// Mitsubishi GX Works2 project: 金达路一号停车场洗车机   PLC: FX3U/FX3UC

PROGRAM MAIN
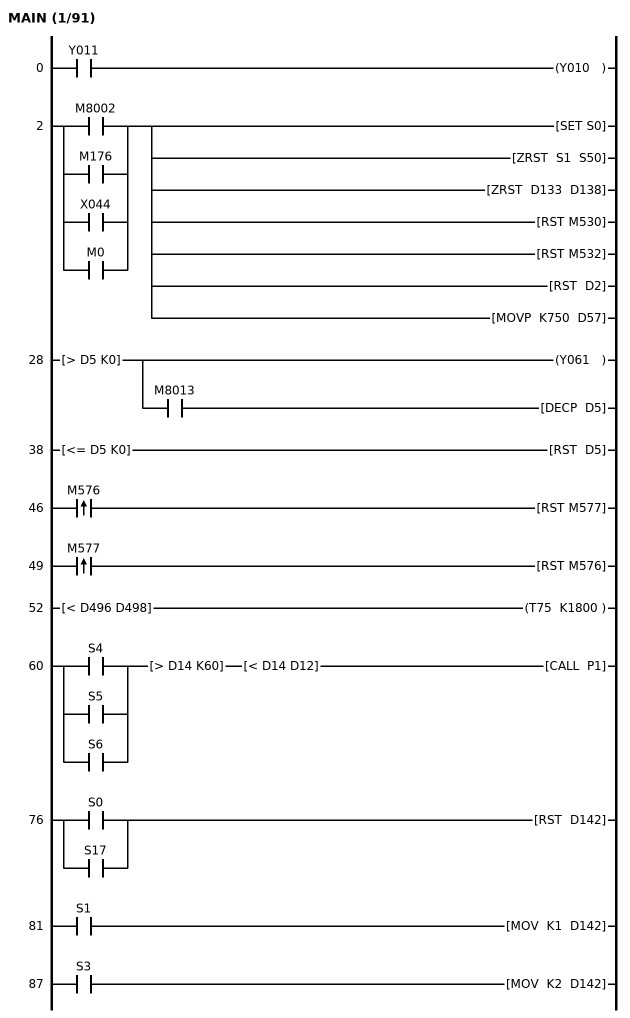
0     LD      Y011
      OUT     Y010
2     LD      M8002
      OR      M176
      OR      X044
      OR      M0
      SET     S0
      ZRST    S1 S50
      ZRST    D133 D138
      RST     M530
      RST     M532
      RST     D2
      MOVP    K750 D57
28    LD>     D5 K0
      OUT     Y061
      AND     M8013
      DECP    D5
38    LD<=    D5 K0
      RST     D5
46    LDP     M576
      RST     M577
49    LDP     M577
      RST     M576
52    LD<     D496 D498
      OUT     T75 K1800
60    LD      S4
      OR      S5
      OR      S6
      AND>    D14 K60
      AND<    D14 D12
      CALL    P1
76    LD      S0
      OR      S17
      RST     D142
81    LD      S1
      MOV     K1 D142
87    LD      S3
      MOV     K2 D142
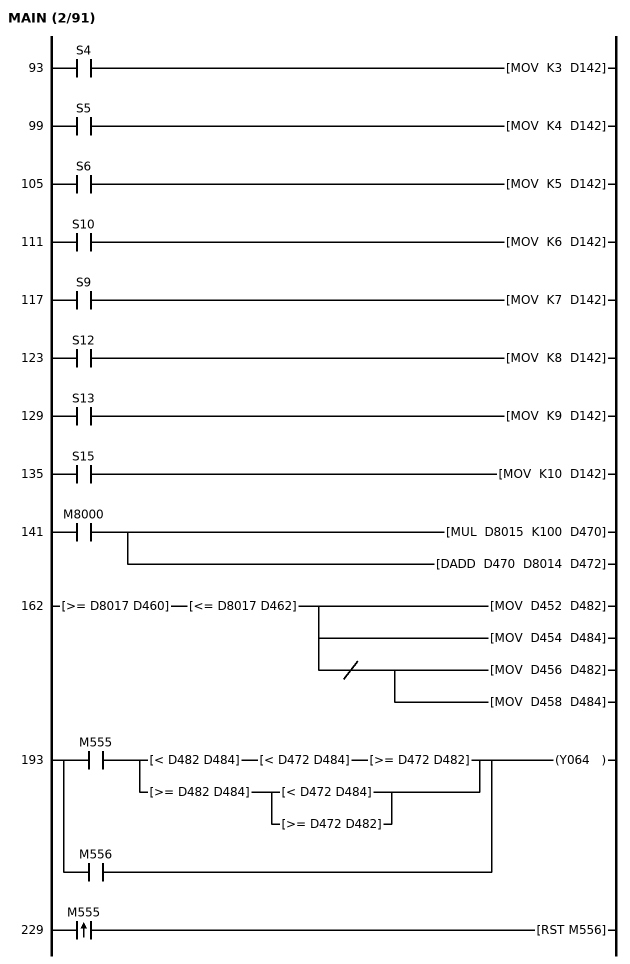
93    LD      S4
      MOV     K3 D142
99    LD      S5
      MOV     K4 D142
105   LD      S6
      MOV     K5 D142
111   LD      S10
      MOV     K6 D142
117   LD      S9
      MOV     K7 D142
123   LD      S12
      MOV     K8 D142
129   LD      S13
      MOV     K9 D142
135   LD      S15
      MOV     K10 D142
141   LD      M8000
      MUL     D8015 K100 D470
      DADD    D470 D8014 D472
162   LD>=    D8017 D460
      AND<=   D8017 D462
      MOV     D452 D482
      MOV     D454 D484
      INV
      MOV     D456 D482
      MOV     D458 D484
193   LD      M555
      LD<     D482 D484
      AND<    D472 D484
      AND>=   D472 D482
      LD>=    D482 D484
      LD<     D472 D484
      OR>=    D472 D482
      ANB
      ORB
      ANB
      OR      M556
      OUT     Y064
229   LDP     M555
      RST     M556
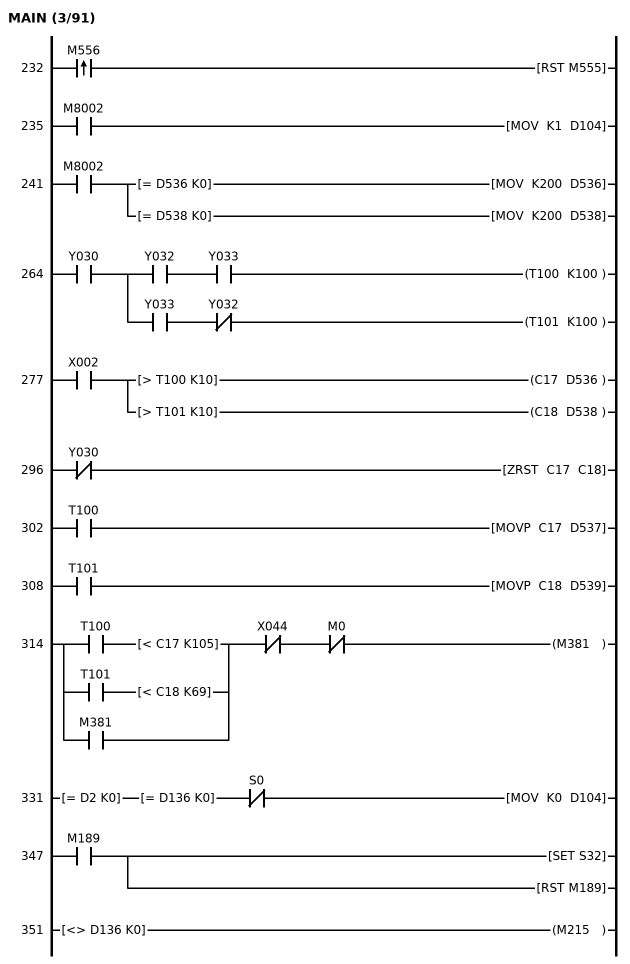
232   LDP     M556
      RST     M555
235   LD      M8002
      MOV     K1 D104
241   LD      M8002
      MPS
      AND=    D536 K0
      MOV     K200 D536
      MPP
      AND=    D538 K0
      MOV     K200 D538
264   LD      Y030
      MPS
      AND     Y032
      AND     Y033
      OUT     T100 K100
      MPP
      AND     Y033
      ANI     Y032
      OUT     T101 K100
277   LD      X002
      MPS
      AND>    T100 K10
      OUT     C17 D536
      MPP
      AND>    T101 K10
      OUT     C18 D538
296   LDI     Y030
      ZRST    C17 C18
302   LD      T100
      MOVP    C17 D537
308   LD      T101
      MOVP    C18 D539
314   LD      T100
      AND<    C17 K105
      LD      T101
      AND<    C18 K69
      ORB
      OR      M381
      ANI     X044
      ANI     M0
      OUT     M381
331   LD=     D2 K0
      AND=    D136 K0
      ANI     S0
      MOV     K0 D104
347   LD      M189
      SET     S32
      RST     M189
351   LD<>    D136 K0
      OUT     M215
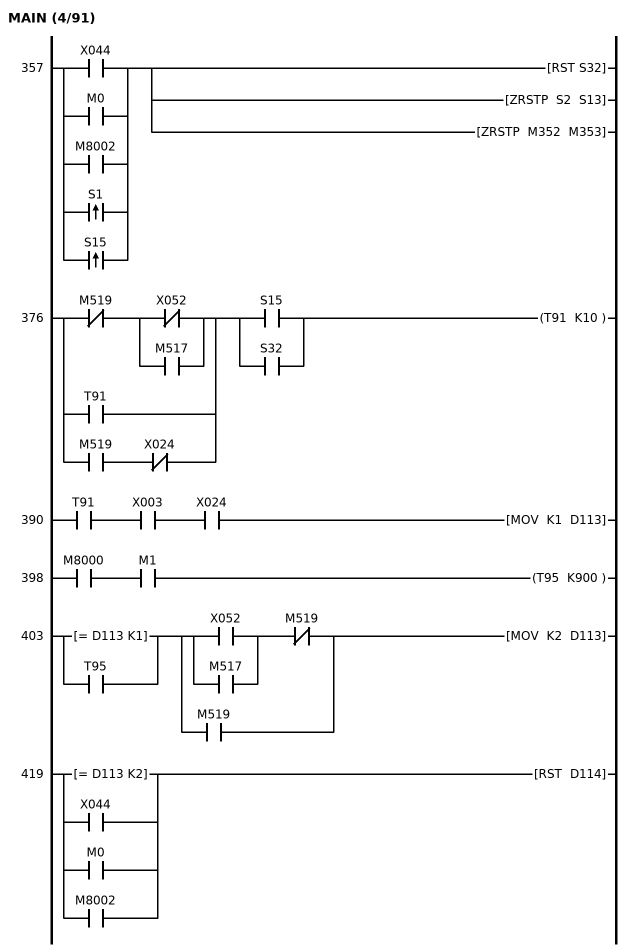
357   LD      X044
      OR      M0
      OR      M8002
      ORP     S1
      ORP     S15
      RST     S32
      ZRSTP   S2 S13
      ZRSTP   M352 M353
376   LDI     M519
      LDI     X052
      OR      M517
      ANB
      OR      T91
      LD      M519
      ANI     X024
      ORB
      LD      S15
      OR      S32
      ANB
      OUT     T91 K10
390   LD      T91
      AND     X003
      AND     X024
      MOV     K1 D113
398   LD      M8000
      AND     M1
      OUT     T95 K900
403   LD=     D113 K1
      OR      T95
      LD      X052
      OR      M517
      ANI     M519
      OR      M519
      ANB
      MOV     K2 D113
419   LD=     D113 K2
      OR      X044
      OR      M0
      OR      M8002
      RST     D114
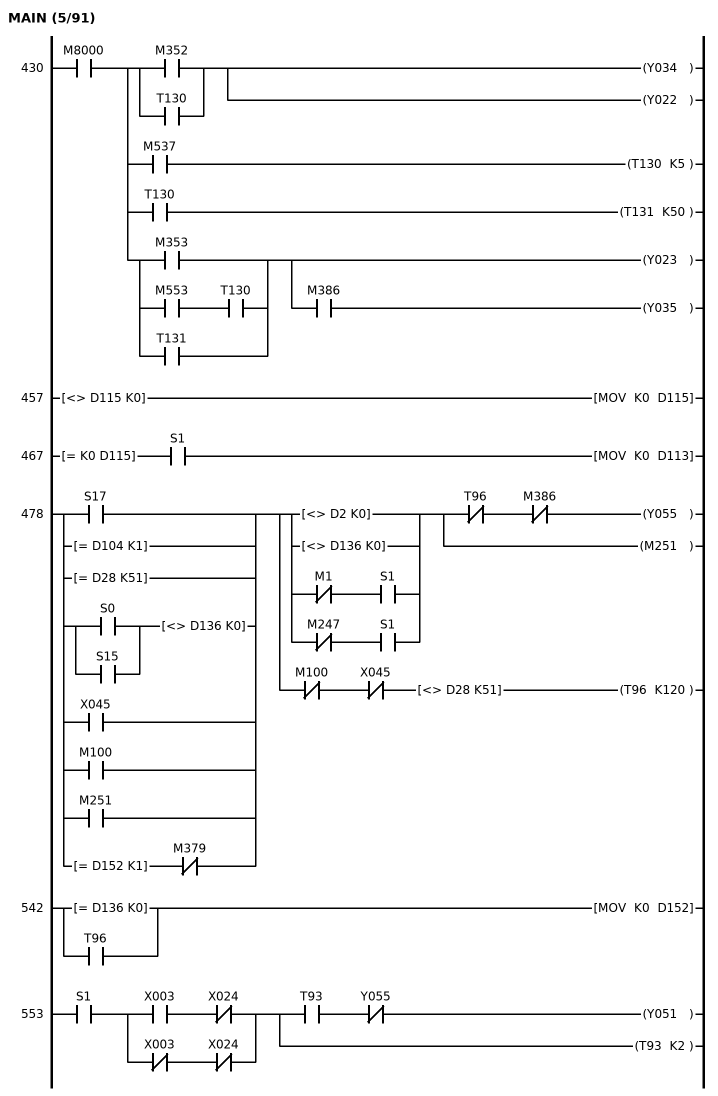
430   LD      M8000
      MPS
      LD      M352
      OR      T130
      ANB
      OUT     Y034
      OUT     Y022
      MRD
      AND     M537
      OUT     T130 K5
      MRD
      AND     T130
      OUT     T131 K50
      MPP
      LD      M353
      LD      M553
      AND     T130
      ORB
      OR      T131
      ANB
      OUT     Y023
      AND     M386
      OUT     Y035
457   LD<>    D115 K0
      MOV     K0 D115
467   LD=     K0 D115
      AND     S1
      MOV     K0 D113
478   LD      S17
      OR=     D104 K1
      OR=     D28 K51
      LD      S0
      OR      S15
      AND<>   D136 K0
      ORB
      OR      X045
      OR      M100
      OR      M251
      LD=     D152 K1
      ANI     M379
      ORB
      MPS
      LD<>    D2 K0
      OR<>    D136 K0
      LDI     M1
      AND     S1
      ORB
      LDI     M247
      AND     S1
      ORB
      ANB
      MPS
      ANI     T96
      ANI     M386
      OUT     Y055
      MPP
      OUT     M251
      MPP
      ANI     M100
      ANI     X045
      AND<>   D28 K51
      OUT     T96 K120
542   LD=     D136 K0
      OR      T96
      MOV     K0 D152
553   LD      S1
      LD      X003
      ANI     X024
      LDI     X003
      ANI     X024
      ORB
      ANB
      MPS
      AND     T93
      ANI     Y055
      OUT     Y051
      MPP
      OUT     T93 K2
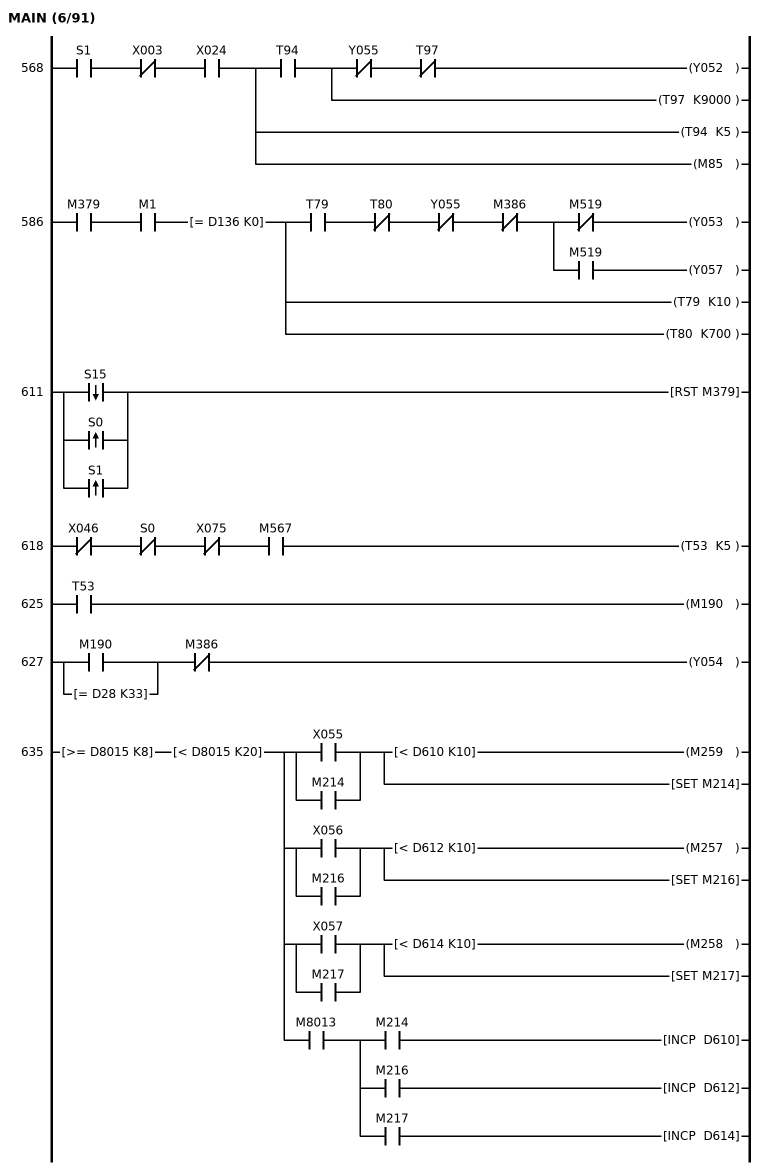
568   LD      S1
      ANI     X003
      AND     X024
      MPS
      AND     T94
      MPS
      ANI     Y055
      ANI     T97
      OUT     Y052
      MPP
      OUT     T97 K9000
      MPP
      OUT     T94 K5
      OUT     M85
586   LD      M379
      AND     M1
      AND=    D136 K0
      MPS
      AND     T79
      ANI     T80
      ANI     Y055
      ANI     M386
      MPS
      ANI     M519
      OUT     Y053
      MPP
      AND     M519
      OUT     Y057
      MPP
      OUT     T79 K10
      OUT     T80 K700
611   LDF     S15
      ORP     S0
      ORP     S1
      RST     M379
618   LDI     X046
      ANI     S0
      ANI     X075
      AND     M567
      OUT     T53 K5
625   LD      T53
      OUT     M190
627   LD      M190
      OR=     D28 K33
      ANI     M386
      OUT     Y054
635   LD>=    D8015 K8
      AND<    D8015 K20
      MPS
      LD      X055
      OR      M214
      ANB
      MPS
      AND<    D610 K10
      OUT     M259
      MPP
      SET     M214
      MRD
      LD      X056
      OR      M216
      ANB
      MPS
      AND<    D612 K10
      OUT     M257
      MPP
      SET     M216
      MRD
      LD      X057
      OR      M217
      ANB
      MPS
      AND<    D614 K10
      OUT     M258
      MPP
      SET     M217
      MPP
      AND     M8013
      MPS
      AND     M214
      INCP    D610
      MRD
      AND     M216
      INCP    D612
      MPP
      AND     M217
      INCP    D614
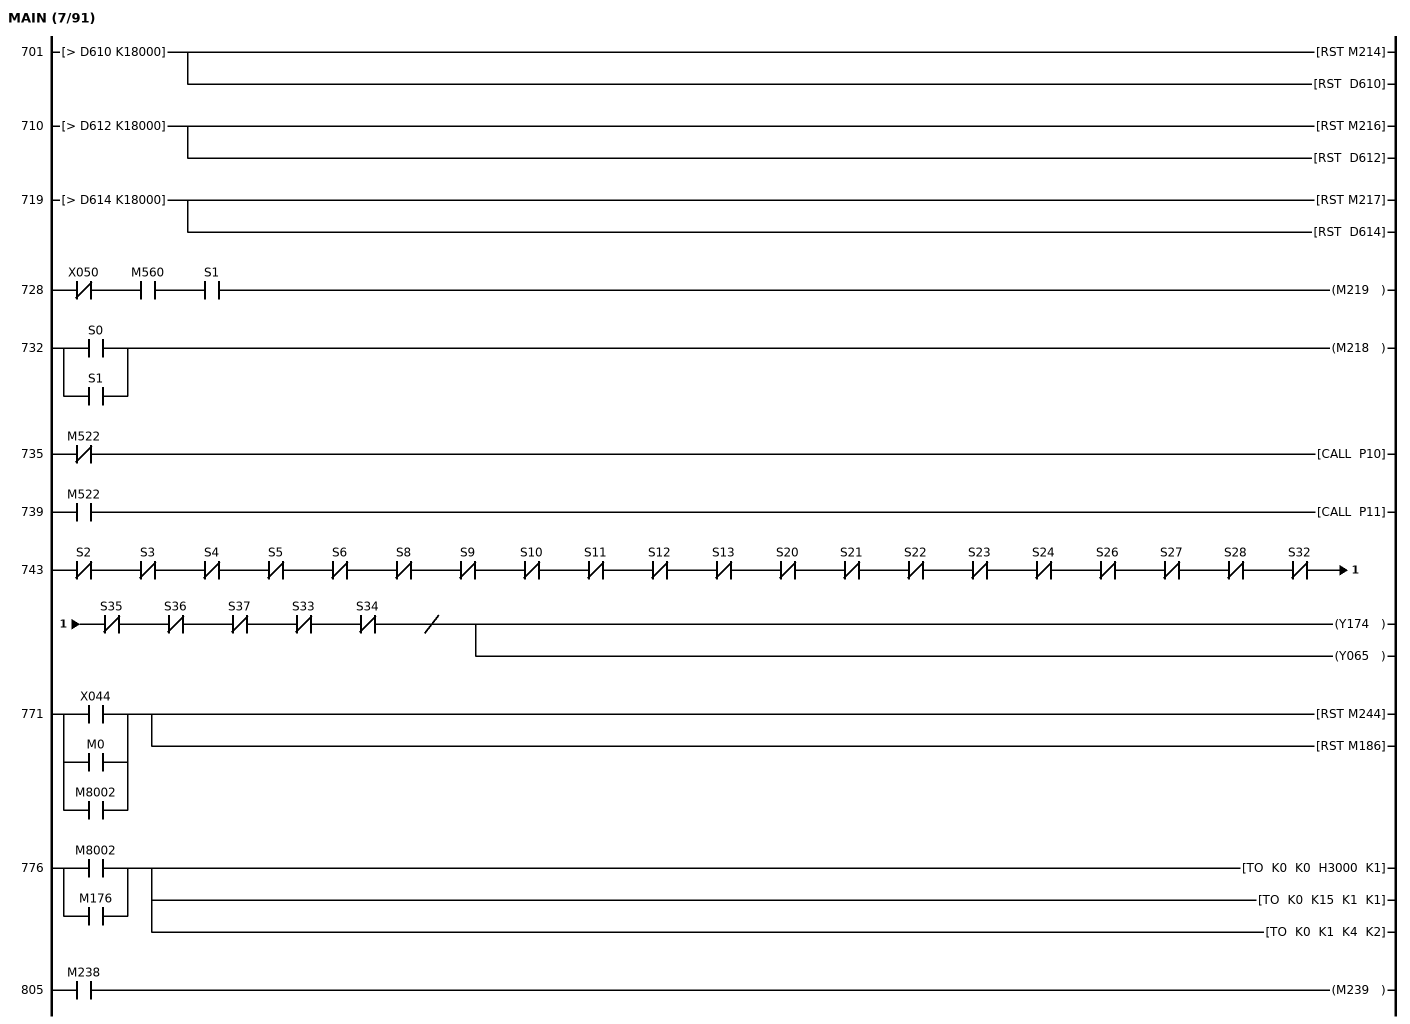
701   LD>     D610 K18000
      RST     M214
      RST     D610
710   LD>     D612 K18000
      RST     M216
      RST     D612
719   LD>     D614 K18000
      RST     M217
      RST     D614
728   LDI     X050
      AND     M560
      AND     S1
      OUT     M219
732   LD      S0
      OR      S1
      OUT     M218
735   LDI     M522
      CALL    P10
739   LD      M522
      CALL    P11
743   LDI     S2
      ANI     S3
      ANI     S4
      ANI     S5
      ANI     S6
      ANI     S8
      ANI     S9
      ANI     S10
      ANI     S11
      ANI     S12
      ANI     S13
      ANI     S20
      ANI     S21
      ANI     S22
      ANI     S23
      ANI     S24
      ANI     S26
      ANI     S27
      ANI     S28
      ANI     S32
      ANI     S35
      ANI     S36
      ANI     S37
      ANI     S33
      ANI     S34
      INV
      OUT     Y174
      OUT     Y065
771   LD      X044
      OR      M0
      OR      M8002
      RST     M244
      RST     M186
776   LD      M8002
      OR      M176
      TO      K0 K0 H3000 K1
      TO      K0 K15 K1 K1
      TO      K0 K1 K4 K2
805   LD      M238
      OUT     M239
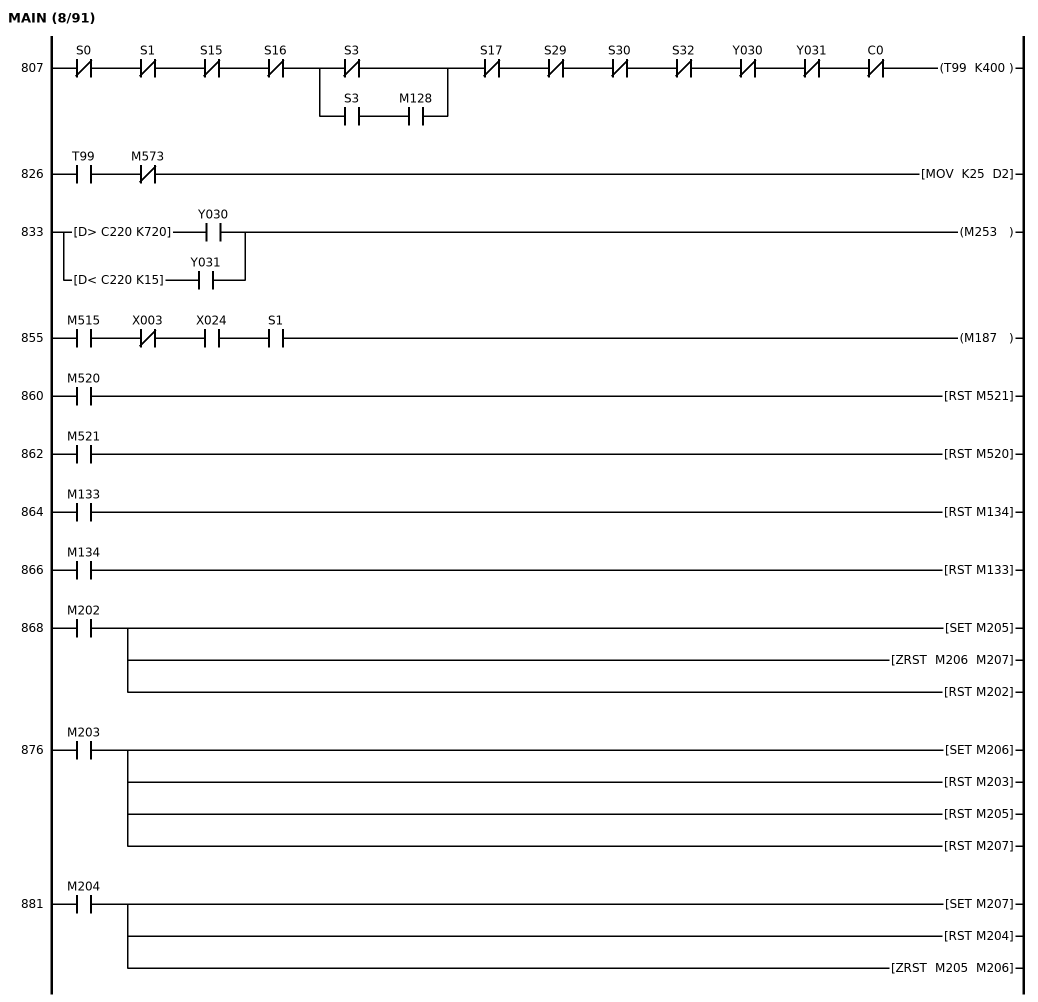
807   LDI     S0
      ANI     S1
      ANI     S15
      ANI     S16
      LDI     S3
      LD      S3
      AND     M128
      ORB
      ANB
      ANI     S17
      ANI     S29
      ANI     S30
      ANI     S32
      ANI     Y030
      ANI     Y031
      ANI     C0
      OUT     T99 K400
826   LD      T99
      ANI     M573
      MOV     K25 D2
833   LDD>    C220 K720
      AND     Y030
      LDD<    C220 K15
      AND     Y031
      ORB
      OUT     M253
855   LD      M515
      ANI     X003
      AND     X024
      AND     S1
      OUT     M187
860   LD      M520
      RST     M521
862   LD      M521
      RST     M520
864   LD      M133
      RST     M134
866   LD      M134
      RST     M133
868   LD      M202
      SET     M205
      ZRST    M206 M207
      RST     M202
876   LD      M203
      SET     M206
      RST     M203
      RST     M205
      RST     M207
881   LD      M204
      SET     M207
      RST     M204
      ZRST    M205 M206
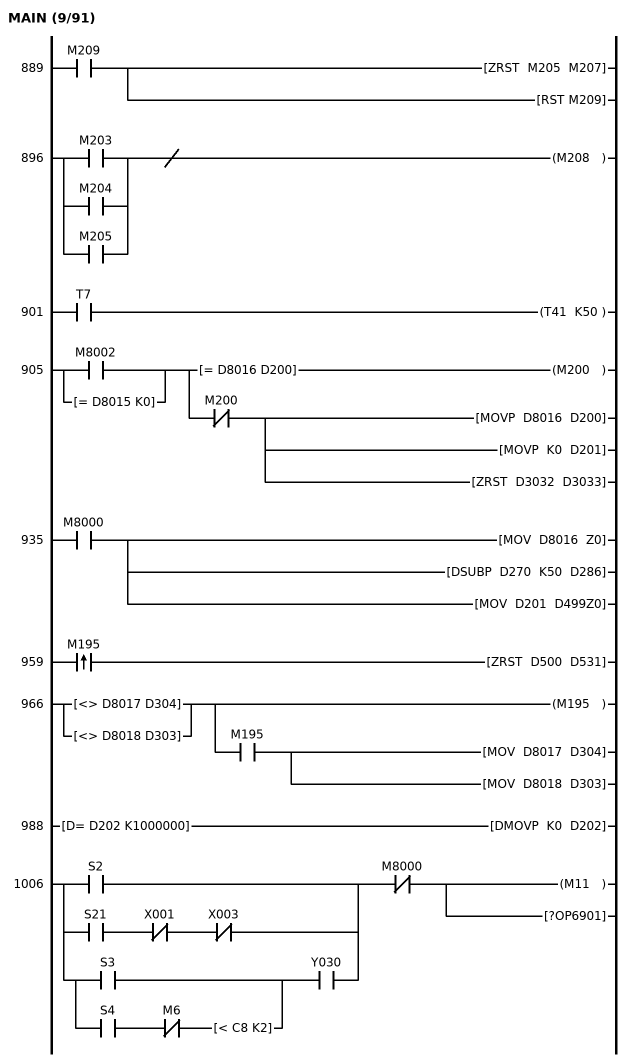
889   LD      M209
      ZRST    M205 M207
      RST     M209
896   LD      M203
      OR      M204
      OR      M205
      INV
      OUT     M208
901   LD      T7
      OUT     T41 K50
905   LD      M8002
      OR=     D8015 K0
      MPS
      AND=    D8016 D200
      OUT     M200
      MPP
      ANI     M200
      MOVP    D8016 D200
      MOVP    K0 D201
      ZRST    D3032 D3033
935   LD      M8000
      MOV     D8016 Z0
      DSUBP   D270 K50 D286
      MOV     D201 D499Z0
959   LDP     M195
      ZRST    D500 D531
966   LD<>    D8017 D304
      OR<>    D8018 D303
      OUT     M195
      AND     M195
      MOV     D8017 D304
      MOV     D8018 D303
988   LDD=    D202 K1000000
      DMOVP   K0 D202
1006  LD      S2
      LD      S21
      ANI     X001
      ANI     X003
      ORB
      LD      S3
      LD      S4
      ANI     M6
      AND<    C8 K2
      ORB
      AND     Y030
      ORB
      ANI     M8000
      OUT     M11
      ?OP6901
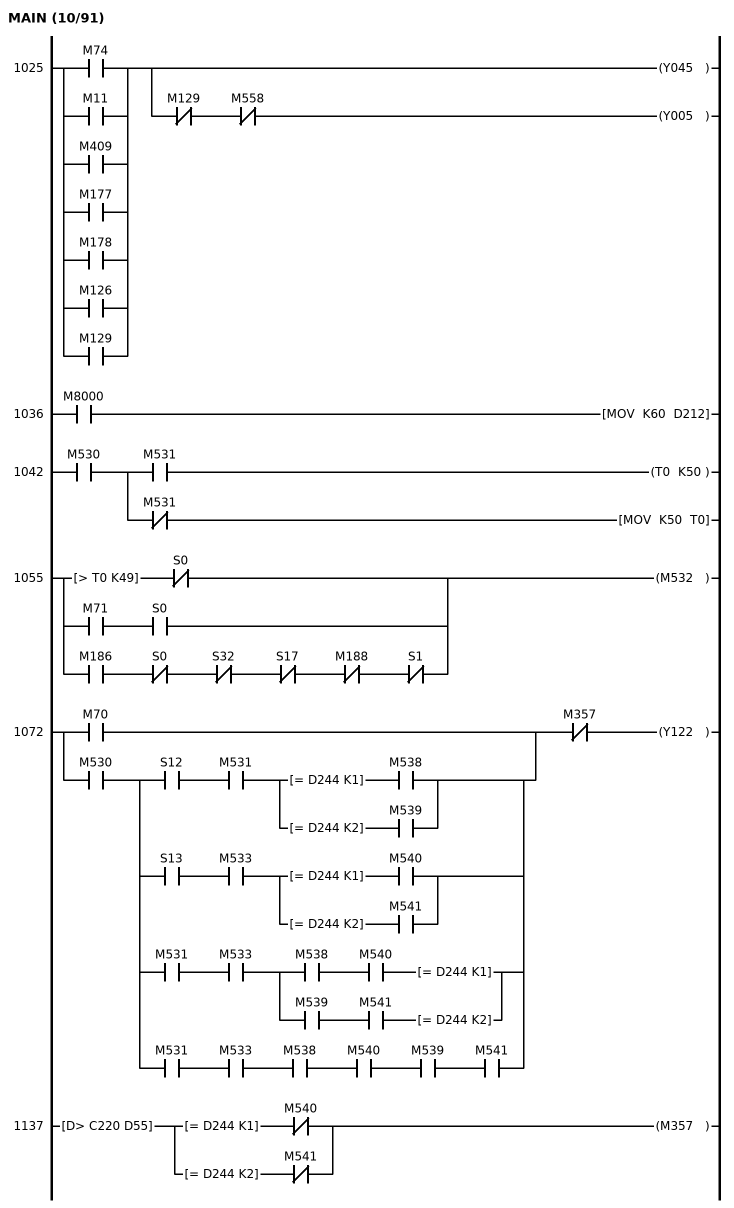
1025  LD      M74
      OR      M11
      OR      M409
      OR      M177
      OR      M178
      OR      M126
      OR      M129
      OUT     Y045
      ANI     M129
      ANI     M558
      OUT     Y005
1036  LD      M8000
      MOV     K60 D212
1042  LD      M530
      MPS
      AND     M531
      OUT     T0 K50
      MPP
      ANI     M531
      MOV     K50 T0
1055  LD>     T0 K49
      ANI     S0
      LD      M71
      AND     S0
      ORB
      LD      M186
      ANI     S0
      ANI     S32
      ANI     S17
      ANI     M188
      ANI     S1
      ORB
      OUT     M532
1072  LD      M70
      LD      M530
      LD      S12
      AND     M531
      LD=     D244 K1
      AND     M538
      LD=     D244 K2
      AND     M539
      ORB
      ANB
      LD      S13
      AND     M533
      LD=     D244 K1
      AND     M540
      LD=     D244 K2
      AND     M541
      ORB
      ANB
      ORB
      LD      M531
      AND     M533
      LD      M538
      AND     M540
      AND=    D244 K1
      LD      M539
      AND     M541
      AND=    D244 K2
      ORB
      ANB
      ORB
      LD      M531
      AND     M533
      AND     M538
      AND     M540
      AND     M539
      AND     M541
      ORB
      ANB
      ORB
      ANI     M357
      OUT     Y122
1137  LDD>    C220 D55
      LD=     D244 K1
      ANI     M540
      LD=     D244 K2
      ANI     M541
      ORB
      ANB
      OUT     M357
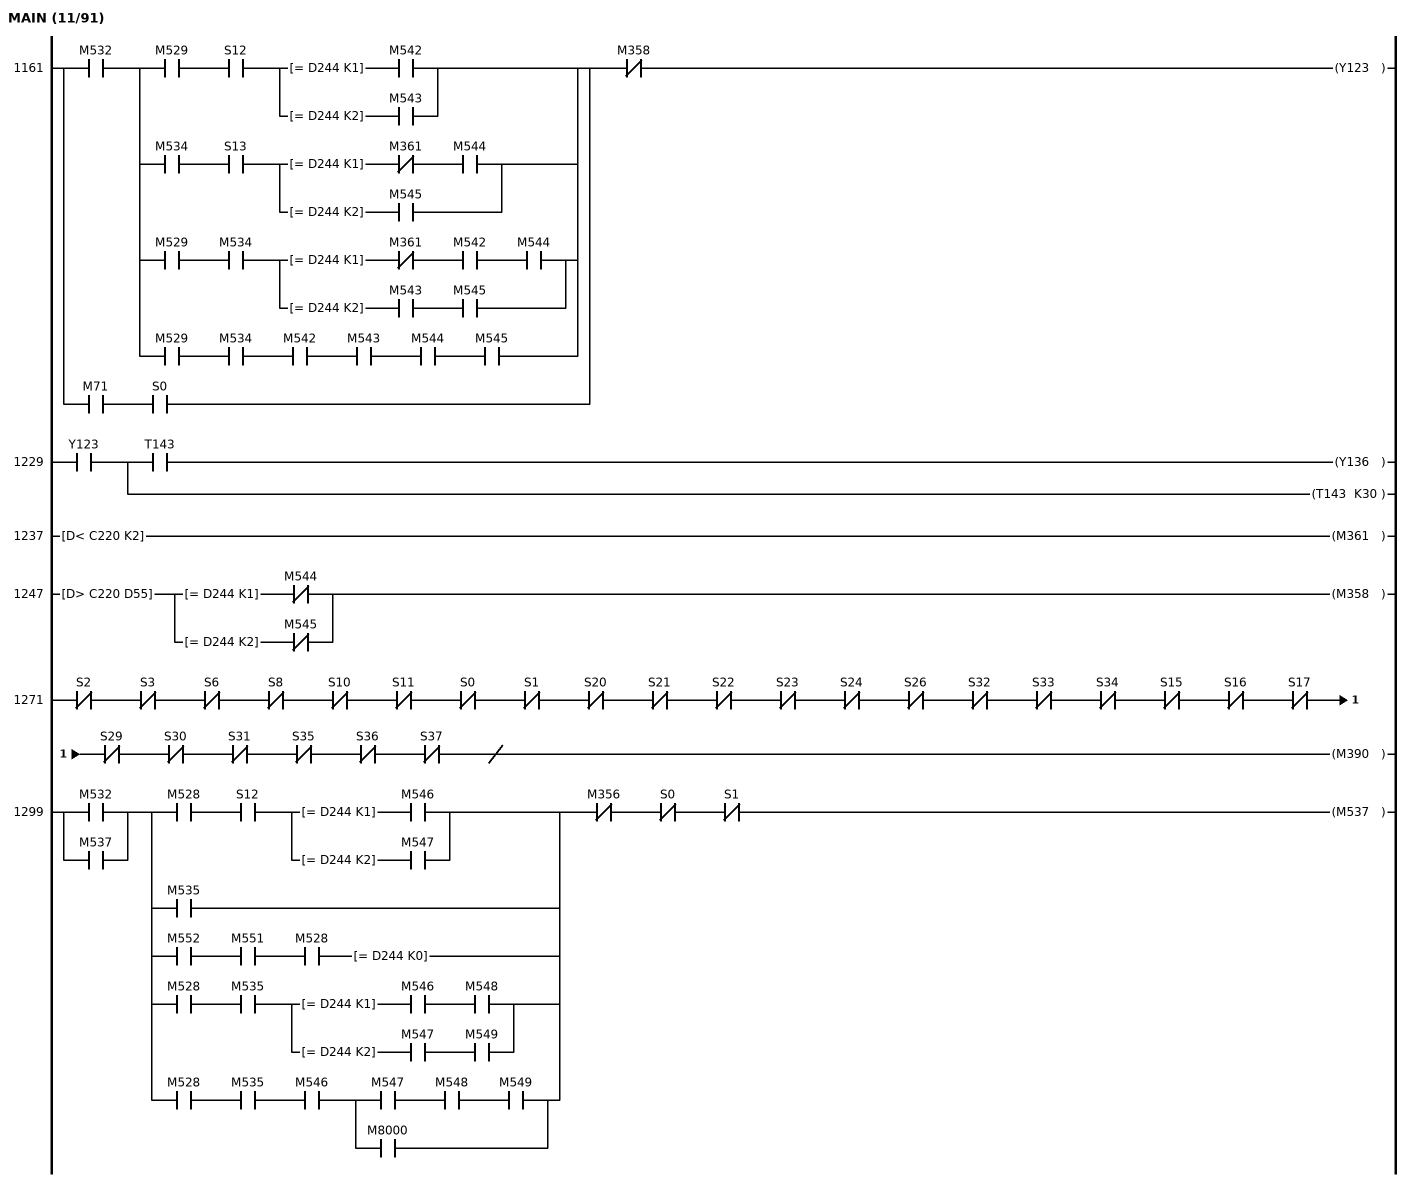
1161  LD      M532
      LD      M529
      AND     S12
      LD=     D244 K1
      AND     M542
      LD=     D244 K2
      AND     M543
      ORB
      ANB
      LD      M534
      AND     S13
      LD=     D244 K1
      ANI     M361
      AND     M544
      LD=     D244 K2
      AND     M545
      ORB
      ANB
      ORB
      LD      M529
      AND     M534
      LD=     D244 K1
      ANI     M361
      AND     M542
      AND     M544
      LD=     D244 K2
      AND     M543
      AND     M545
      ORB
      ANB
      ORB
      LD      M529
      AND     M534
      AND     M542
      AND     M543
      AND     M544
      AND     M545
      ORB
      ANB
      LD      M71
      AND     S0
      ORB
      ANI     M358
      OUT     Y123
1229  LD      Y123
      MPS
      AND     T143
      OUT     Y136
      MPP
      OUT     T143 K30
1237  LDD<    C220 K2
      OUT     M361
1247  LDD>    C220 D55
      LD=     D244 K1
      ANI     M544
      LD=     D244 K2
      ANI     M545
      ORB
      ANB
      OUT     M358
1271  LDI     S2
      ANI     S3
      ANI     S6
      ANI     S8
      ANI     S10
      ANI     S11
      ANI     S0
      ANI     S1
      ANI     S20
      ANI     S21
      ANI     S22
      ANI     S23
      ANI     S24
      ANI     S26
      ANI     S32
      ANI     S33
      ANI     S34
      ANI     S15
      ANI     S16
      ANI     S17
      ANI     S29
      ANI     S30
      ANI     S31
      ANI     S35
      ANI     S36
      ANI     S37
      INV
      OUT     M390
1299  LD      M532
      OR      M537
      LD      M528
      AND     S12
      LD=     D244 K1
      AND     M546
      LD=     D244 K2
      AND     M547
      ORB
      ANB
      OR      M535
      LD      M552
      AND     M551
      AND     M528
      AND=    D244 K0
      ORB
      LD      M528
      AND     M535
      LD=     D244 K1
      AND     M546
      AND     M548
      LD=     D244 K2
      AND     M547
      AND     M549
      ORB
      ANB
      ORB
      LD      M528
      AND     M535
      AND     M546
      LD      M547
      AND     M548
      AND     M549
      OR      M8000
      ANB
      ORB
      ANB
      ANI     M356
      ANI     S0
      ANI     S1
      OUT     M537
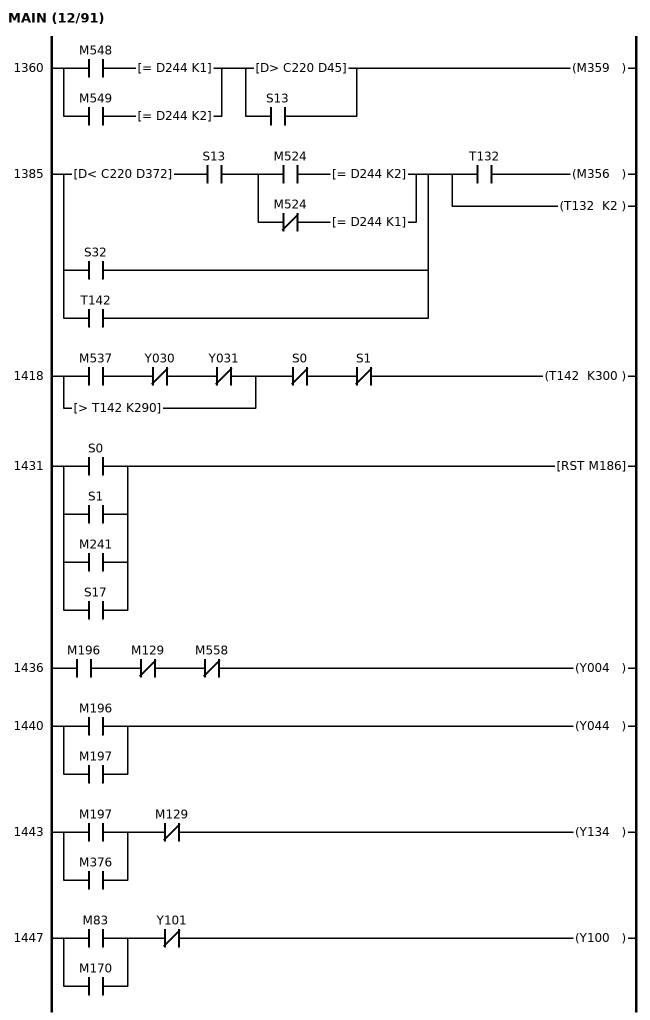
1360  LD      M548
      AND=    D244 K1
      LD      M549
      AND=    D244 K2
      ORB
      LDD>    C220 D45
      OR      S13
      ANB
      OUT     M359
1385  LDD<    C220 D372
      AND     S13
      LD      M524
      AND=    D244 K2
      LDI     M524
      AND=    D244 K1
      ORB
      ANB
      OR      S32
      OR      T142
      MPS
      AND     T132
      OUT     M356
      MPP
      OUT     T132 K2
1418  LD      M537
      ANI     Y030
      ANI     Y031
      OR>     T142 K290
      ANI     S0
      ANI     S1
      OUT     T142 K300
1431  LD      S0
      OR      S1
      OR      M241
      OR      S17
      RST     M186
1436  LD      M196
      ANI     M129
      ANI     M558
      OUT     Y004
1440  LD      M196
      OR      M197
      OUT     Y044
1443  LD      M197
      OR      M376
      ANI     M129
      OUT     Y134
1447  LD      M83
      OR      M170
      ANI     Y101
      OUT     Y100
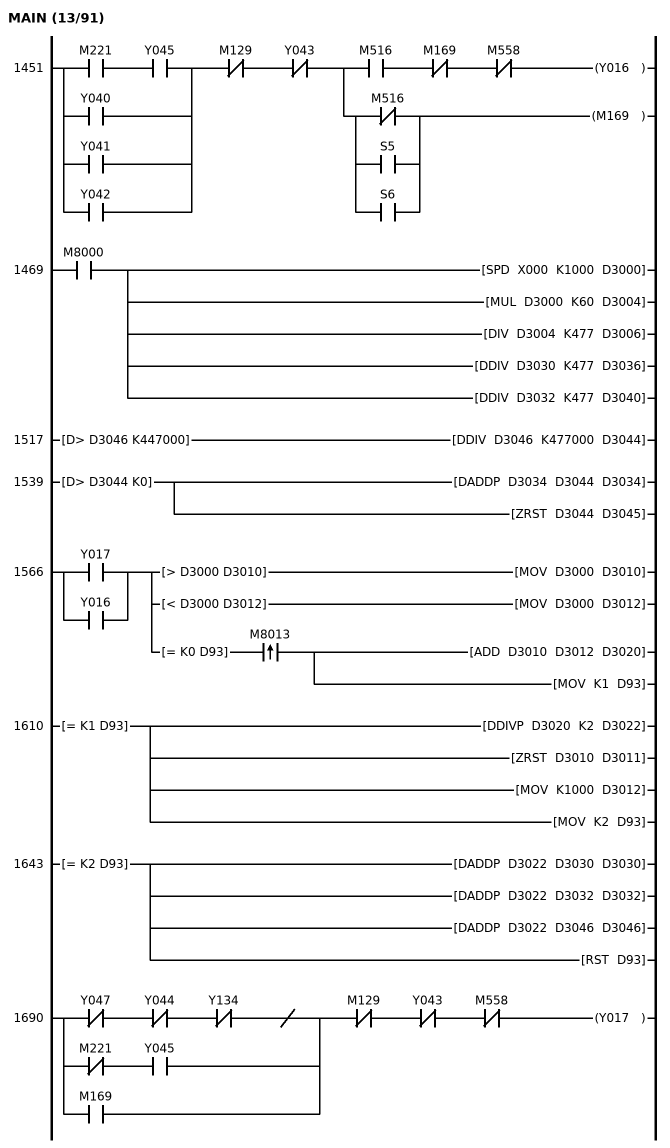
1451  LD      M221
      AND     Y045
      OR      Y040
      OR      Y041
      OR      Y042
      ANI     M129
      ANI     Y043
      MPS
      AND     M516
      ANI     M169
      ANI     M558
      OUT     Y016
      MPP
      LDI     M516
      OR      S5
      OR      S6
      ANB
      OUT     M169
1469  LD      M8000
      SPD     X000 K1000 D3000
      MUL     D3000 K60 D3004
      DIV     D3004 K477 D3006
      DDIV    D3030 K477 D3036
      DDIV    D3032 K477 D3040
1517  LDD>    D3046 K447000
      DDIV    D3046 K477000 D3044
1539  LDD>    D3044 K0
      DADDP   D3034 D3044 D3034
      ZRST    D3044 D3045
1566  LD      Y017
      OR      Y016
      MPS
      AND>    D3000 D3010
      MOV     D3000 D3010
      MRD
      AND<    D3000 D3012
      MOV     D3000 D3012
      MPP
      AND=    K0 D93
      ANDP    M8013
      ADD     D3010 D3012 D3020
      MOV     K1 D93
1610  LD=     K1 D93
      DDIVP   D3020 K2 D3022
      ZRST    D3010 D3011
      MOV     K1000 D3012
      MOV     K2 D93
1643  LD=     K2 D93
      DADDP   D3022 D3030 D3030
      DADDP   D3022 D3032 D3032
      DADDP   D3022 D3046 D3046
      RST     D93
1690  LDI     Y047
      ANI     Y044
      ANI     Y134
      INV
      LDI     M221
      AND     Y045
      ORB
      OR      M169
      ANI     M129
      ANI     Y043
      ANI     M558
      OUT     Y017
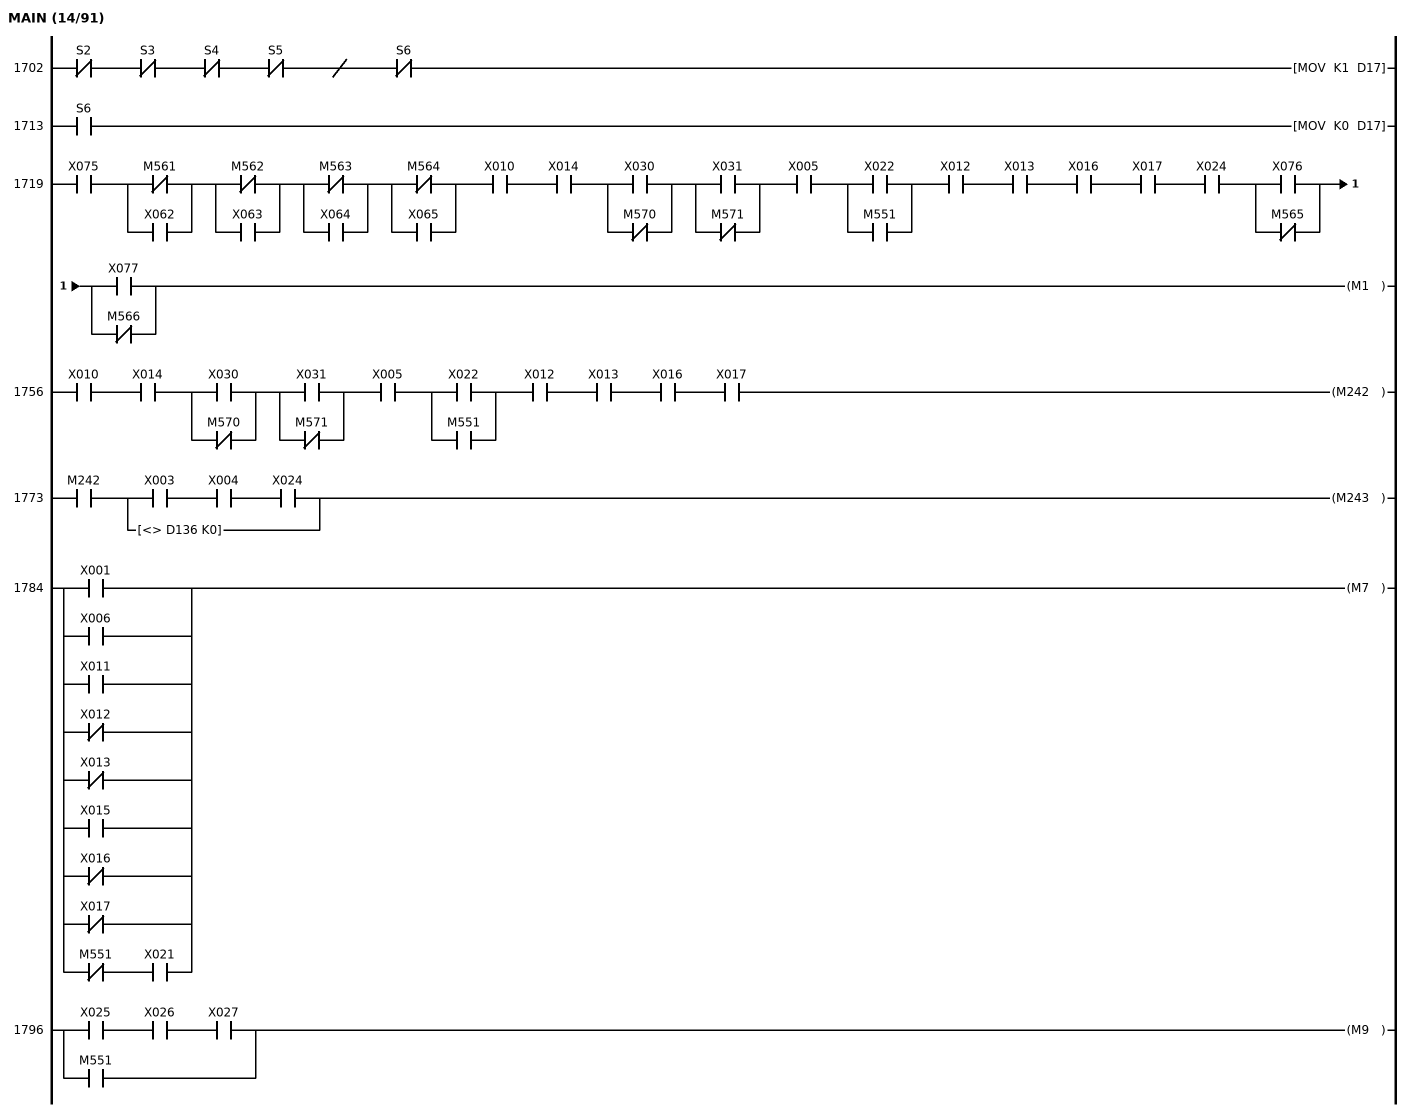
1702  LDI     S2
      ANI     S3
      ANI     S4
      ANI     S5
      INV
      ANI     S6
      MOV     K1 D17
1713  LD      S6
      MOV     K0 D17
1719  LD      X075
      LDI     M561
      OR      X062
      ANB
      LDI     M562
      OR      X063
      ANB
      LDI     M563
      OR      X064
      ANB
      LDI     M564
      OR      X065
      ANB
      AND     X010
      AND     X014
      LD      X030
      ORI     M570
      ANB
      LD      X031
      ORI     M571
      ANB
      AND     X005
      LD      X022
      OR      M551
      ANB
      AND     X012
      AND     X013
      AND     X016
      AND     X017
      AND     X024
      LD      X076
      ORI     M565
      ANB
      LD      X077
      ORI     M566
      ANB
      OUT     M1
1756  LD      X010
      AND     X014
      LD      X030
      ORI     M570
      ANB
      LD      X031
      ORI     M571
      ANB
      AND     X005
      LD      X022
      OR      M551
      ANB
      AND     X012
      AND     X013
      AND     X016
      AND     X017
      OUT     M242
1773  LD      M242
      LD      X003
      AND     X004
      AND     X024
      OR<>    D136 K0
      ANB
      OUT     M243
1784  LD      X001
      OR      X006
      OR      X011
      ORI     X012
      ORI     X013
      OR      X015
      ORI     X016
      ORI     X017
      LDI     M551
      AND     X021
      ORB
      OUT     M7
1796  LD      X025
      AND     X026
      AND     X027
      OR      M551
      OUT     M9
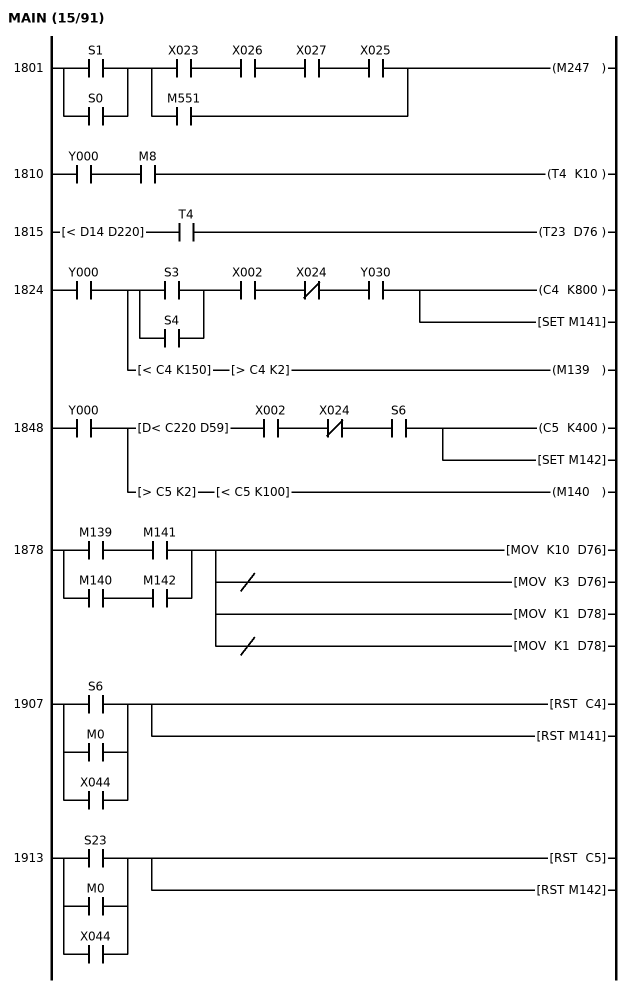
1801  LD      S1
      OR      S0
      LD      X023
      AND     X026
      AND     X027
      AND     X025
      OR      M551
      ANB
      OUT     M247
1810  LD      Y000
      AND     M8
      OUT     T4 K10
1815  LD<     D14 D220
      AND     T4
      OUT     T23 D76
1824  LD      Y000
      MPS
      LD      S3
      OR      S4
      ANB
      AND     X002
      ANI     X024
      AND     Y030
      OUT     C4 K800
      SET     M141
      MPP
      AND<    C4 K150
      AND>    C4 K2
      OUT     M139
1848  LD      Y000
      MPS
      ANDD<   C220 D59
      AND     X002
      ANI     X024
      AND     S6
      OUT     C5 K400
      SET     M142
      MPP
      AND>    C5 K2
      AND<    C5 K100
      OUT     M140
1878  LD      M139
      AND     M141
      LD      M140
      AND     M142
      ORB
      MOV     K10 D76
      MPS
      INV
      MOV     K3 D76
      MPP
      MOV     K1 D78
      INV
      MOV     K1 D78
1907  LD      S6
      OR      M0
      OR      X044
      RST     C4
      RST     M141
1913  LD      S23
      OR      M0
      OR      X044
      RST     C5
      RST     M142
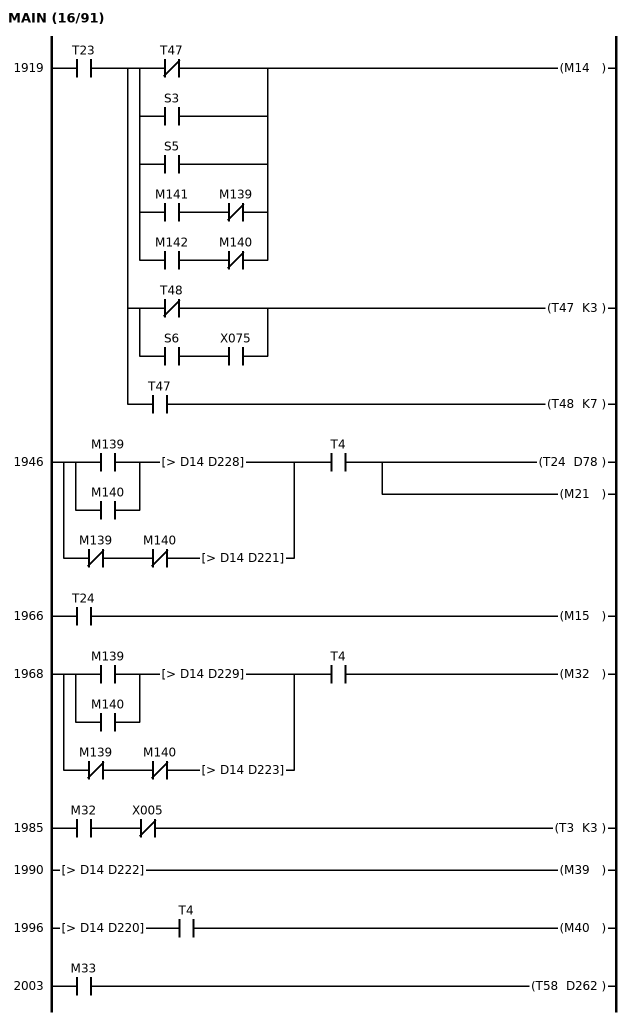
1919  LD      T23
      MPS
      LDI     T47
      OR      S3
      OR      S5
      LD      M141
      ANI     M139
      ORB
      LD      M142
      ANI     M140
      ORB
      ANB
      OUT     M14
      MRD
      LDI     T48
      LD      S6
      AND     X075
      ORB
      ANB
      OUT     T47 K3
      MPP
      AND     T47
      OUT     T48 K7
1946  LD      M139
      OR      M140
      AND>    D14 D228
      LDI     M139
      ANI     M140
      AND>    D14 D221
      ORB
      AND     T4
      OUT     T24 D78
      OUT     M21
1966  LD      T24
      OUT     M15
1968  LD      M139
      OR      M140
      AND>    D14 D229
      LDI     M139
      ANI     M140
      AND>    D14 D223
      ORB
      AND     T4
      OUT     M32
1985  LD      M32
      ANI     X005
      OUT     T3 K3
1990  LD>     D14 D222
      OUT     M39
1996  LD>     D14 D220
      AND     T4
      OUT     M40
2003  LD      M33
      OUT     T58 D262
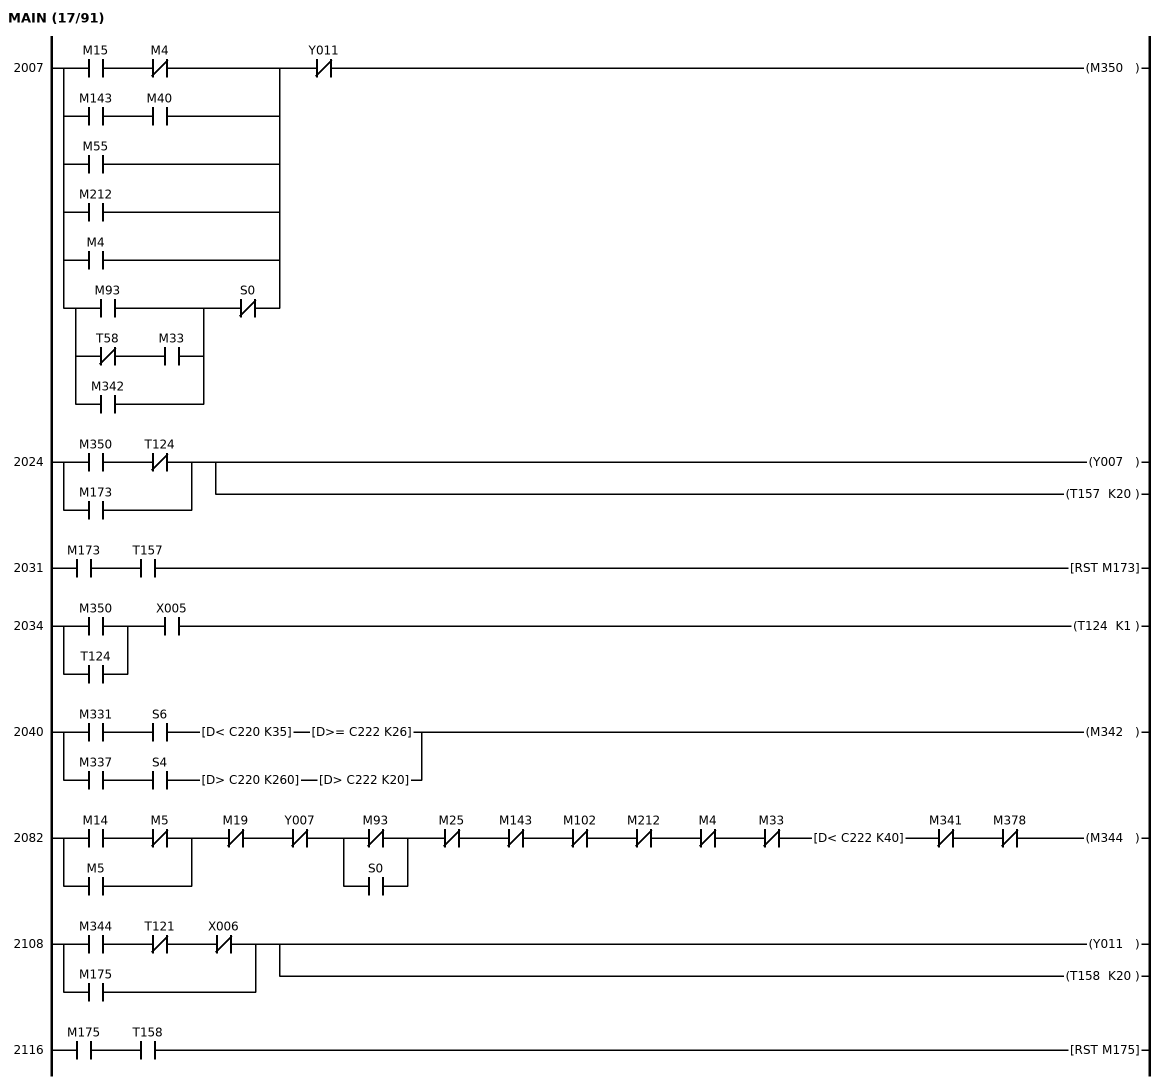
2007  LD      M15
      ANI     M4
      LD      M143
      AND     M40
      ORB
      OR      M55
      OR      M212
      OR      M4
      LD      M93
      LDI     T58
      AND     M33
      ORB
      OR      M342
      ANI     S0
      ORB
      ANI     Y011
      OUT     M350
2024  LD      M350
      ANI     T124
      OR      M173
      OUT     Y007
      OUT     T157 K20
2031  LD      M173
      AND     T157
      RST     M173
2034  LD      M350
      OR      T124
      AND     X005
      OUT     T124 K1
2040  LD      M331
      AND     S6
      ANDD<   C220 K35
      ANDD>=  C222 K26
      LD      M337
      AND     S4
      ANDD>   C220 K260
      ANDD>   C222 K20
      ORB
      OUT     M342
2082  LD      M14
      ANI     M5
      OR      M5
      ANI     M19
      ANI     Y007
      LDI     M93
      OR      S0
      ANB
      ANI     M25
      ANI     M143
      ANI     M102
      ANI     M212
      ANI     M4
      ANI     M33
      ANDD<   C222 K40
      ANI     M341
      ANI     M378
      OUT     M344
2108  LD      M344
      ANI     T121
      ANI     X006
      OR      M175
      OUT     Y011
      OUT     T158 K20
2116  LD      M175
      AND     T158
      RST     M175
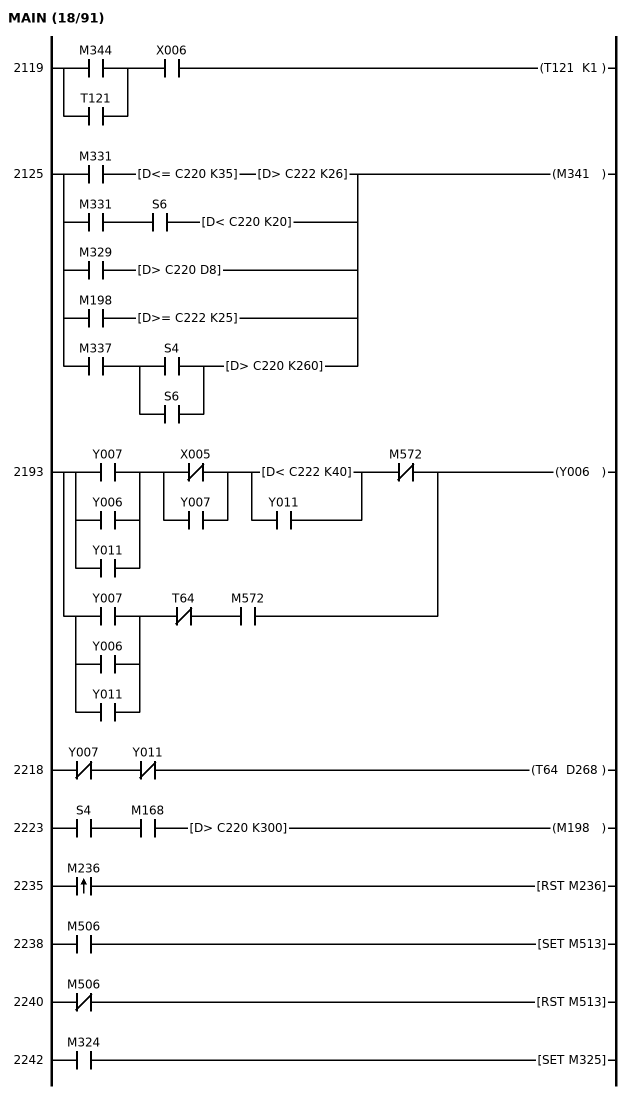
2119  LD      M344
      OR      T121
      AND     X006
      OUT     T121 K1
2125  LD      M331
      ANDD<=  C220 K35
      ANDD>   C222 K26
      LD      M331
      AND     S6
      ANDD<   C220 K20
      ORB
      LD      M329
      ANDD>   C220 D8
      ORB
      LD      M198
      ANDD>=  C222 K25
      ORB
      LD      M337
      LD      S4
      OR      S6
      ANB
      ANDD>   C220 K260
      ORB
      OUT     M341
2193  LD      Y007
      OR      Y006
      OR      Y011
      LDI     X005
      OR      Y007
      ANB
      LDD<    C222 K40
      OR      Y011
      ANB
      ANI     M572
      LD      Y007
      OR      Y006
      OR      Y011
      ANI     T64
      AND     M572
      ORB
      OUT     Y006
2218  LDI     Y007
      ANI     Y011
      OUT     T64 D268
2223  LD      S4
      AND     M168
      ANDD>   C220 K300
      OUT     M198
2235  LDP     M236
      RST     M236
2238  LD      M506
      SET     M513
2240  LDI     M506
      RST     M513
2242  LD      M324
      SET     M325
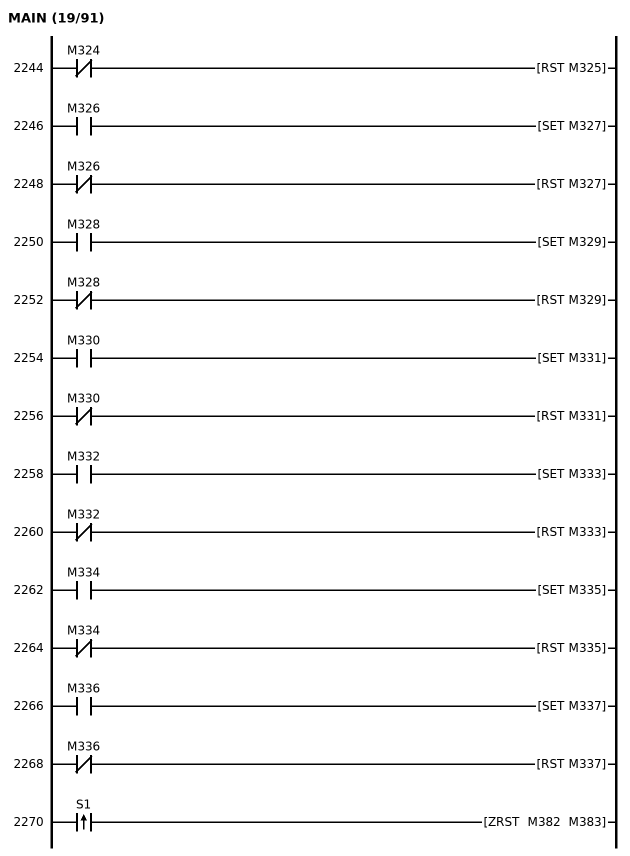
2244  LDI     M324
      RST     M325
2246  LD      M326
      SET     M327
2248  LDI     M326
      RST     M327
2250  LD      M328
      SET     M329
2252  LDI     M328
      RST     M329
2254  LD      M330
      SET     M331
2256  LDI     M330
      RST     M331
2258  LD      M332
      SET     M333
2260  LDI     M332
      RST     M333
2262  LD      M334
      SET     M335
2264  LDI     M334
      RST     M335
2266  LD      M336
      SET     M337
2268  LDI     M336
      RST     M337
2270  LDP     S1
      ZRST    M382 M383
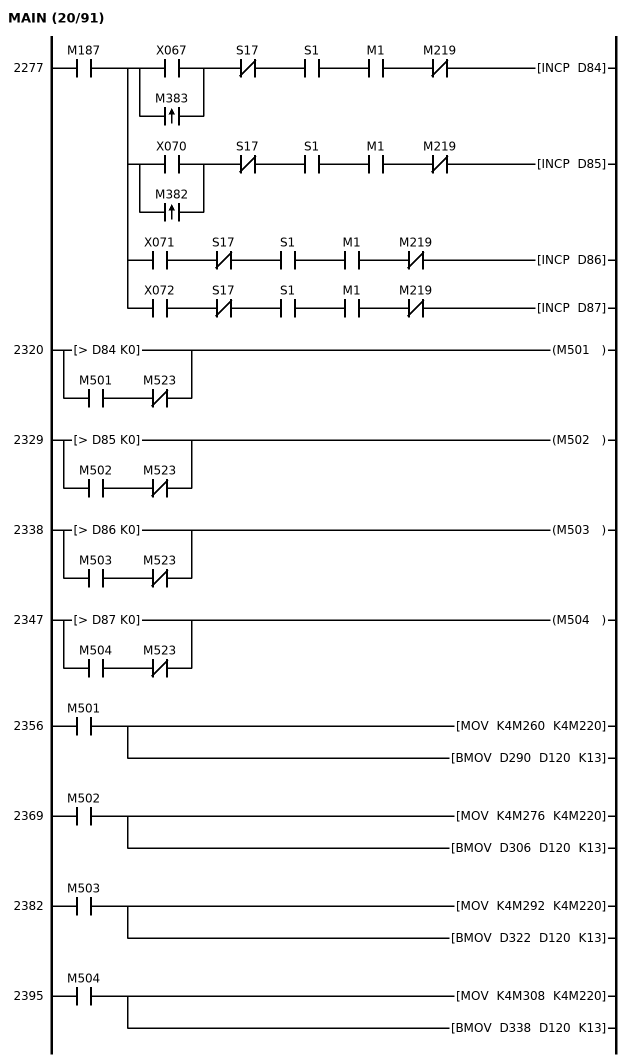
2277  LD      M187
      MPS
      LD      X067
      ORP     M383
      ANB
      ANI     S17
      AND     S1
      AND     M1
      ANI     M219
      INCP    D84
      MRD
      LD      X070
      ORP     M382
      ANB
      ANI     S17
      AND     S1
      AND     M1
      ANI     M219
      INCP    D85
      MRD
      AND     X071
      ANI     S17
      AND     S1
      AND     M1
      ANI     M219
      INCP    D86
      MPP
      AND     X072
      ANI     S17
      AND     S1
      AND     M1
      ANI     M219
      INCP    D87
2320  LD>     D84 K0
      LD      M501
      ANI     M523
      ORB
      OUT     M501
2329  LD>     D85 K0
      LD      M502
      ANI     M523
      ORB
      OUT     M502
2338  LD>     D86 K0
      LD      M503
      ANI     M523
      ORB
      OUT     M503
2347  LD>     D87 K0
      LD      M504
      ANI     M523
      ORB
      OUT     M504
2356  LD      M501
      MOV     K4M260 K4M220
      BMOV    D290 D120 K13
2369  LD      M502
      MOV     K4M276 K4M220
      BMOV    D306 D120 K13
2382  LD      M503
      MOV     K4M292 K4M220
      BMOV    D322 D120 K13
2395  LD      M504
      MOV     K4M308 K4M220
      BMOV    D338 D120 K13
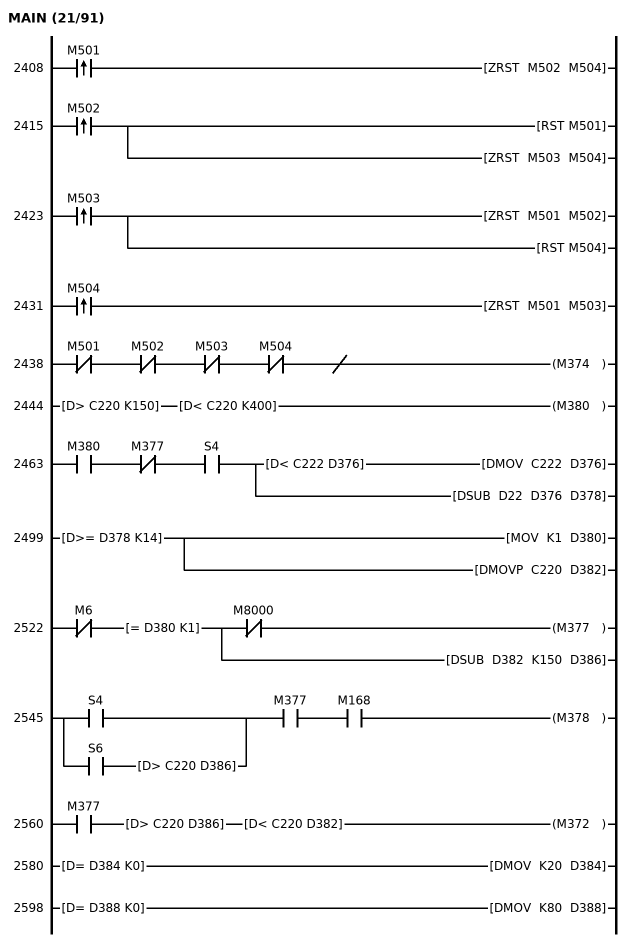
2408  LDP     M501
      ZRST    M502 M504
2415  LDP     M502
      RST     M501
      ZRST    M503 M504
2423  LDP     M503
      ZRST    M501 M502
      RST     M504
2431  LDP     M504
      ZRST    M501 M503
2438  LDI     M501
      ANI     M502
      ANI     M503
      ANI     M504
      INV
      OUT     M374
2444  LDD>    C220 K150
      ANDD<   C220 K400
      OUT     M380
2463  LD      M380
      ANI     M377
      AND     S4
      MPS
      ANDD<   C222 D376
      DMOV    C222 D376
      MPP
      DSUB    D22 D376 D378
2499  LDD>=   D378 K14
      MOV     K1 D380
      DMOVP   C220 D382
2522  LDI     M6
      AND=    D380 K1
      MPS
      ANI     M8000
      OUT     M377
      MPP
      DSUB    D382 K150 D386
2545  LD      S4
      LD      S6
      ANDD>   C220 D386
      ORB
      AND     M377
      AND     M168
      OUT     M378
2560  LD      M377
      ANDD>   C220 D386
      ANDD<   C220 D382
      OUT     M372
2580  LDD=    D384 K0
      DMOV    K20 D384
2598  LDD=    D388 K0
      DMOV    K80 D388
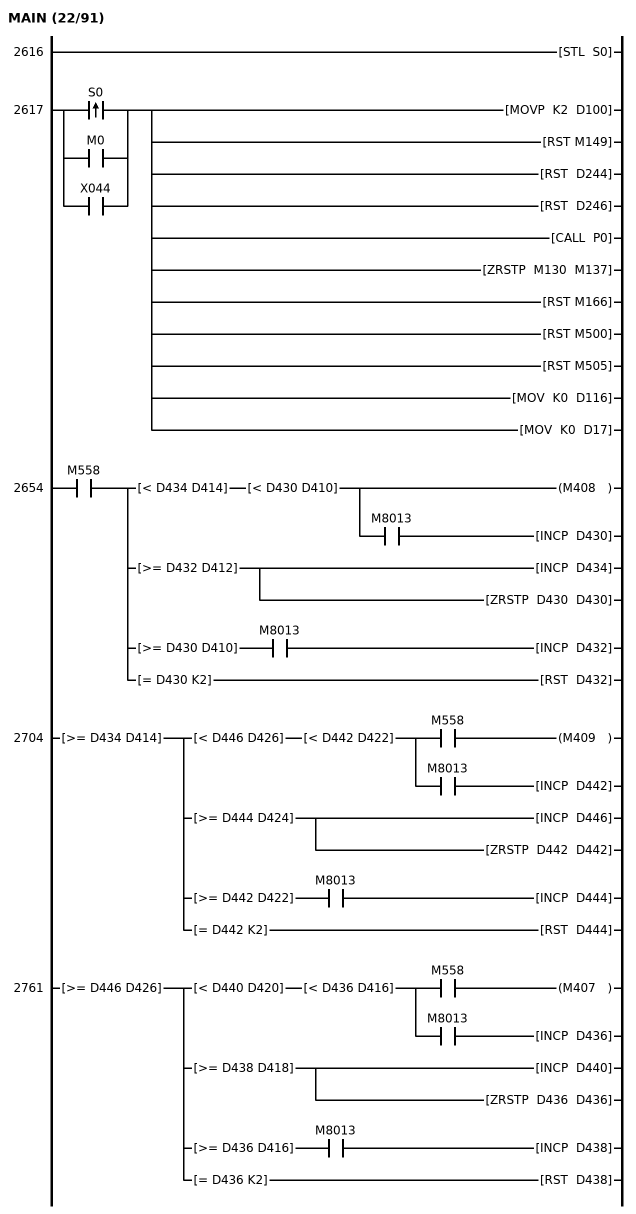
2616  STL     S0
2617  LDP     S0
      OR      M0
      OR      X044
      MOVP    K2 D100
      RST     M149
      RST     D244
      RST     D246
      CALL    P0
      ZRSTP   M130 M137
      RST     M166
      RST     M500
      RST     M505
      MOV     K0 D116
      MOV     K0 D17
2654  LD      M558
      MPS
      AND<    D434 D414
      AND<    D430 D410
      OUT     M408
      AND     M8013
      INCP    D430
      MRD
      AND>=   D432 D412
      INCP    D434
      ZRSTP   D430 D430
      MRD
      AND>=   D430 D410
      AND     M8013
      INCP    D432
      MPP
      AND=    D430 K2
      RST     D432
2704  LD>=    D434 D414
      MPS
      AND<    D446 D426
      AND<    D442 D422
      MPS
      AND     M558
      OUT     M409
      MPP
      AND     M8013
      INCP    D442
      MRD
      AND>=   D444 D424
      INCP    D446
      ZRSTP   D442 D442
      MRD
      AND>=   D442 D422
      AND     M8013
      INCP    D444
      MPP
      AND=    D442 K2
      RST     D444
2761  LD>=    D446 D426
      MPS
      AND<    D440 D420
      AND<    D436 D416
      MPS
      AND     M558
      OUT     M407
      MPP
      AND     M8013
      INCP    D436
      MRD
      AND>=   D438 D418
      INCP    D440
      ZRSTP   D436 D436
      MRD
      AND>=   D436 D416
      AND     M8013
      INCP    D438
      MPP
      AND=    D436 K2
      RST     D438
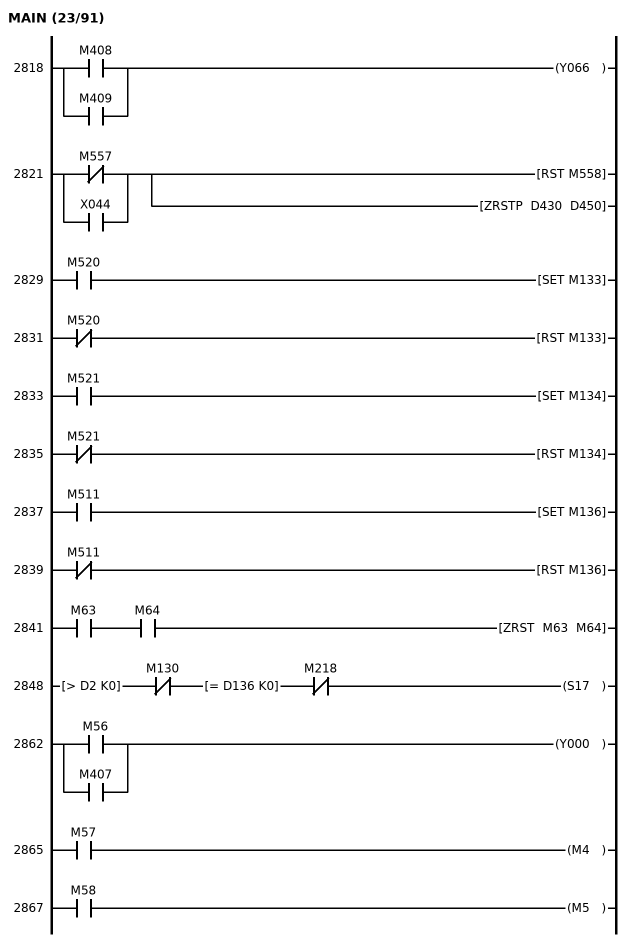
2818  LD      M408
      OR      M409
      OUT     Y066
2821  LDI     M557
      OR      X044
      RST     M558
      ZRSTP   D430 D450
2829  LD      M520
      SET     M133
2831  LDI     M520
      RST     M133
2833  LD      M521
      SET     M134
2835  LDI     M521
      RST     M134
2837  LD      M511
      SET     M136
2839  LDI     M511
      RST     M136
2841  LD      M63
      AND     M64
      ZRST    M63 M64
2848  LD>     D2 K0
      ANI     M130
      AND=    D136 K0
      ANI     M218
      OUT     S17
2862  LD      M56
      OR      M407
      OUT     Y000
2865  LD      M57
      OUT     M4
2867  LD      M58
      OUT     M5
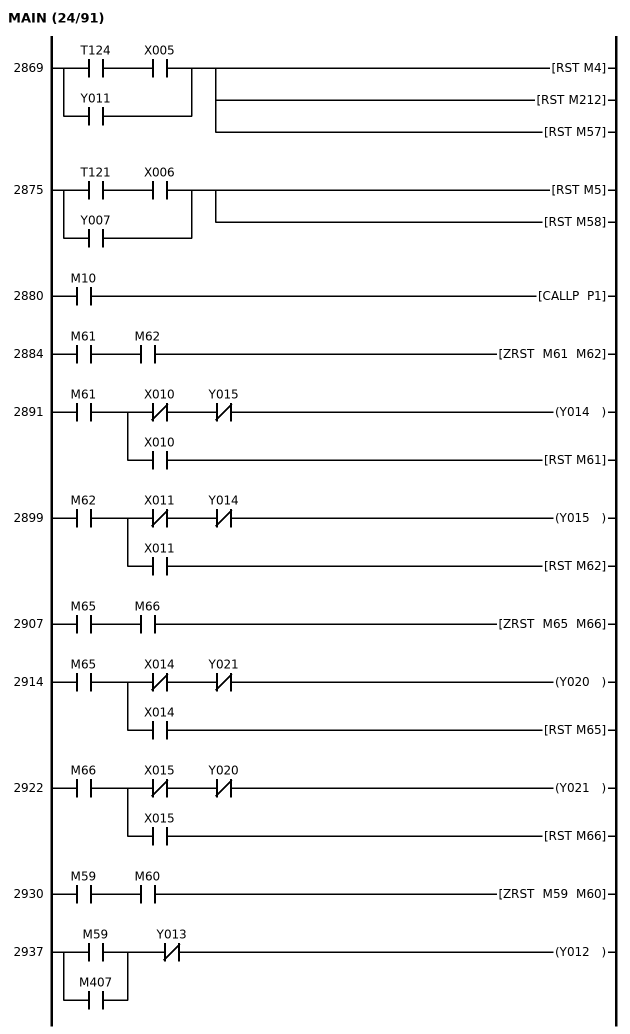
2869  LD      T124
      AND     X005
      OR      Y011
      RST     M4
      RST     M212
      RST     M57
2875  LD      T121
      AND     X006
      OR      Y007
      RST     M5
      RST     M58
2880  LD      M10
      CALLP   P1
2884  LD      M61
      AND     M62
      ZRST    M61 M62
2891  LD      M61
      MPS
      ANI     X010
      ANI     Y015
      OUT     Y014
      MPP
      AND     X010
      RST     M61
2899  LD      M62
      MPS
      ANI     X011
      ANI     Y014
      OUT     Y015
      MPP
      AND     X011
      RST     M62
2907  LD      M65
      AND     M66
      ZRST    M65 M66
2914  LD      M65
      MPS
      ANI     X014
      ANI     Y021
      OUT     Y020
      MPP
      AND     X014
      RST     M65
2922  LD      M66
      MPS
      ANI     X015
      ANI     Y020
      OUT     Y021
      MPP
      AND     X015
      RST     M66
2930  LD      M59
      AND     M60
      ZRST    M59 M60
2937  LD      M59
      OR      M407
      ANI     Y013
      OUT     Y012
